// TIA Portal V21 export
// export: Created 2026-08-21T20:18:54.0096754Z, ExportSetting None, DisplayName Totally Integrated Automation Portal, DisplayVersion V21, DisplayName STEP 7 Professional, DisplayVersion V21, DisplayName STEP 7 Safety, DisplayVersion V21, DisplayName Tech WebApplication, DisplayVersion V21, DisplayName WinCC Basic/Comfort/Advanced, DisplayVersion V21, DisplayName WinCC Professional, DisplayVersion V21, DisplayName WinCC Unified, DisplayVersion V21
FUNCTION_BLOCK "MTPPIDCtrl_Type1"   // FB14, FBD
{ S7_Optimized_Access := 'TRUE' }
// stored: MemoryReserve 100, SetENOAutomatically false
   VAR_INPUT
      from_Actor { ExternalAccessible := 'False'; ExternalVisible := 'False'; ExternalWritable := 'False'} : "StruCm";
      SP_Ext { ExternalAccessible := 'False'; ExternalVisible := 'False'; ExternalWritable := 'False'} : Real;
      Service_Occupied { ExternalAccessible := 'False'; ExternalVisible := 'False'; ExternalWritable := 'False'} : Bool;
      Cmd_Auto { ExternalAccessible := 'False'; ExternalVisible := 'False'; ExternalWritable := 'False'} : Bool;
      Cmd_Man { ExternalAccessible := 'False'; ExternalVisible := 'False'; ExternalWritable := 'False'} : Bool;
      Cmd_SPExt { ExternalAccessible := 'False'; ExternalVisible := 'False'; ExternalWritable := 'False'} : Bool;
      Cmd_SPInt { ExternalAccessible := 'False'; ExternalVisible := 'False'; ExternalWritable := 'False'} : Bool;
      PV { ExternalAccessible := 'False'; ExternalVisible := 'False'; ExternalWritable := 'False'} : Word;
      PV_QB { ExternalAccessible := 'False'; ExternalVisible := 'False'; ExternalWritable := 'False'} : Bool := true;
      PV_Unit { ExternalAccessible := 'False'; ExternalVisible := 'False'; ExternalWritable := 'False'} : Int := 1342;
      Intlk04_In01 { ExternalAccessible := 'False'; ExternalVisible := 'False'; ExternalWritable := 'False'} : "DigVal";
      Intlk04_InvIn01 { ExternalAccessible := 'False'; ExternalVisible := 'False'; ExternalWritable := 'False'} : Bool;
      Intlk04_In1String : String;
      Intlk04_In02 { ExternalAccessible := 'False'; ExternalVisible := 'False'; ExternalWritable := 'False'} : "DigVal";
      Intlk04_InvIn02 { ExternalAccessible := 'False'; ExternalVisible := 'False'; ExternalWritable := 'False'} : Bool;
      Intlk04_In2String : String;
      Intlk04_In03 { ExternalAccessible := 'False'; ExternalVisible := 'False'; ExternalWritable := 'False'} : "DigVal";
      Intlk04_InvIn03 { ExternalAccessible := 'False'; ExternalVisible := 'False'; ExternalWritable := 'False'} : Bool;
      Intlk04_In3String : String;
      Intlk04_In04 { ExternalAccessible := 'False'; ExternalVisible := 'False'; ExternalWritable := 'False'} : "DigVal";
      Intlk04_InvIn04 { ExternalAccessible := 'False'; ExternalVisible := 'False'; ExternalWritable := 'False'} : Bool;
      Intlk04_In4String : String;
   END_VAR
   VAR_OUTPUT
      to_Actor { ExternalAccessible := 'False'; ExternalVisible := 'False'; ExternalWritable := 'False'} : "StruCm";
      Occupied { ExternalAccessible := 'False'; ExternalVisible := 'False'; ExternalWritable := 'False'} : Bool;   // Occupied by a Service procedure
      AutAct { ExternalAccessible := 'False'; ExternalVisible := 'False'; ExternalWritable := 'False'} : Bool;
      ManAct { ExternalAccessible := 'False'; ExternalVisible := 'False'; ExternalWritable := 'False'} : Bool;
      SP_ExtAct { ExternalAccessible := 'False'; ExternalVisible := 'False'; ExternalWritable := 'False'} : Bool;
      GrpErr { ExternalAccessible := 'False'; ExternalVisible := 'False'; ExternalWritable := 'False'} : Bool;
      PV_AH_Act { ExternalAccessible := 'False'; ExternalVisible := 'False'; ExternalWritable := 'False'} : Bool;
      PV_WH_Act { ExternalAccessible := 'False'; ExternalVisible := 'False'; ExternalWritable := 'False'} : Bool;
      PV_WL_Act { ExternalAccessible := 'False'; ExternalVisible := 'False'; ExternalWritable := 'False'} : Bool;
      PV_AL_Act { ExternalAccessible := 'False'; ExternalVisible := 'False'; ExternalWritable := 'False'} : Bool;
   END_VAR
   VAR
      AnIn_IDB { ExternalAccessible := 'False'; ExternalVisible := 'False'; ExternalWritable := 'False'} : "AnIn";
      Intlk04_IDB : "Intlk04";
      PIDConL_IDB { S7_SetPoint := 'True'} : "PIDConL";
      MTPPIDCtrl_IDB { ExternalVisible := 'False'; S7_SetPoint := 'True'} : "MTPPIDCtrl";
   END_VAR
   VAR_TEMP
      Intlock : "DigVal";
      PV_Out : "AnaVal";
      ScaleOut : "ScaVal";
      BadOut : "DigVal";
      CSF_NOP : "DigVal";
   END_VAR
   // Intlk04_In01.Value := true;
   // Intlk04_In02.Value := true;
   // Intlk04_In03.Value := true;
   // Intlk04_In04.Value := true;
BEGIN

REGION Network 1: Mod switch
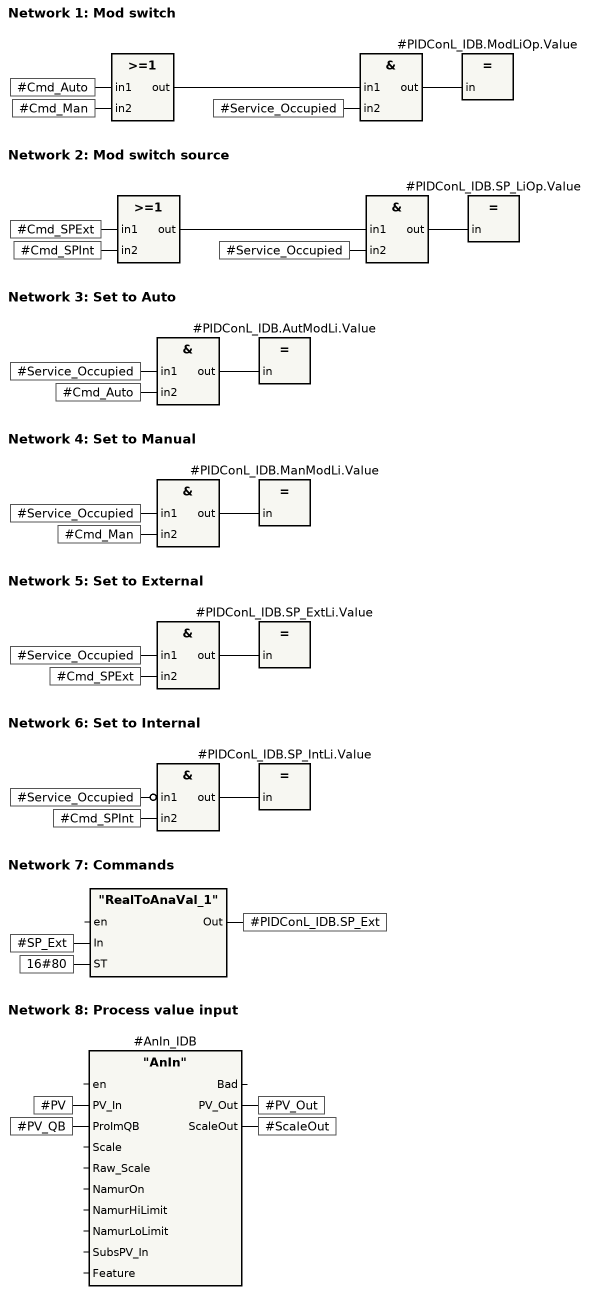
   #PIDConL_IDB.ModLiOp.Value := (#Cmd_Auto OR #Cmd_Man) AND #Service_Occupied;
END_REGION

REGION Network 2: Mod switch source
   #PIDConL_IDB.SP_LiOp.Value := (#Cmd_SPExt OR #Cmd_SPInt) AND #Service_Occupied;
END_REGION

REGION Network 3: Set to Auto
   #PIDConL_IDB.AutModLi.Value := #Service_Occupied AND #Cmd_Auto;
END_REGION

REGION Network 4: Set to Manual
   #PIDConL_IDB.ManModLi.Value := #Service_Occupied AND #Cmd_Man;
END_REGION

REGION Network 5: Set to External
   #PIDConL_IDB.SP_ExtLi.Value := #Service_Occupied AND #Cmd_SPExt;
END_REGION

REGION Network 6: Set to Internal
   #PIDConL_IDB.SP_IntLi.Value := NOT #Service_Occupied AND #Cmd_SPInt;
END_REGION

REGION Network 7: Commands
   "RealToAnaVal_1"(In := #SP_Ext, ST := 16#80, Out => #PIDConL_IDB.SP_Ext);
END_REGION

REGION Network 8: Process value input
   #AnIn_IDB(PV_In := #PV, ProImQB := #PV_QB, PV_Out => #PV_Out, ScaleOut => #ScaleOut);   // "AnIn"
END_REGION

REGION Network 9: CSF
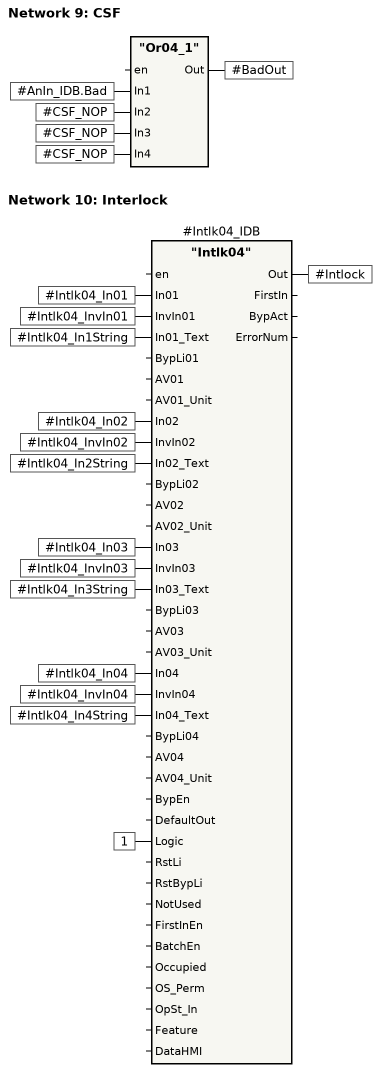
   "Or04_1"(In1 := #AnIn_IDB.Bad, In2 := #CSF_NOP, In3 := #CSF_NOP, In4 := #CSF_NOP, Out => #BadOut);
END_REGION

REGION Network 10: Interlock
   #Intlk04_IDB(In01 := #Intlk04_In01,   // "Intlk04"
                InvIn01 := #Intlk04_InvIn01,
                In01_Text := #Intlk04_In1String,
                In02 := #Intlk04_In02,
                InvIn02 := #Intlk04_InvIn02,
                In02_Text := #Intlk04_In2String,
                In03 := #Intlk04_In03,
                InvIn03 := #Intlk04_InvIn03,
                In03_Text := #Intlk04_In3String,
                In04 := #Intlk04_In04,
                InvIn04 := #Intlk04_InvIn04,
                In04_Text := #Intlk04_In4String,
                Logic := 1,
                Out => #Intlock);
END_REGION

REGION Network 11: PIDCtrL / PIDConL
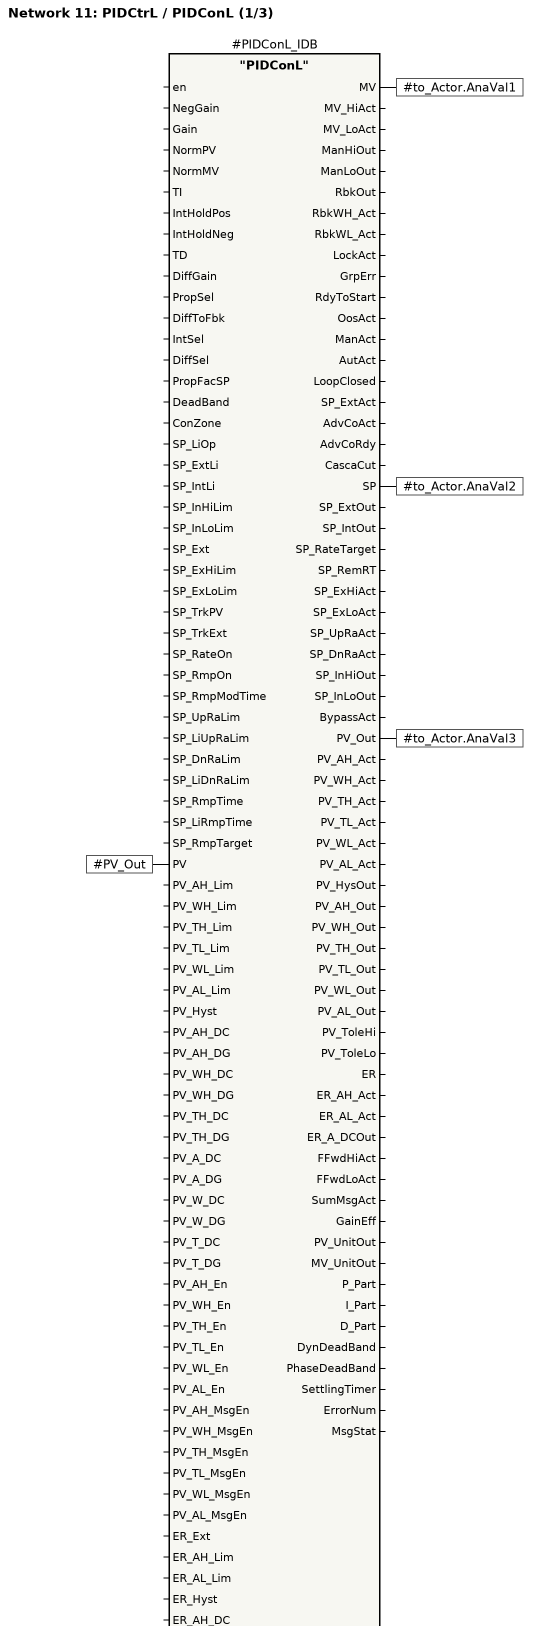
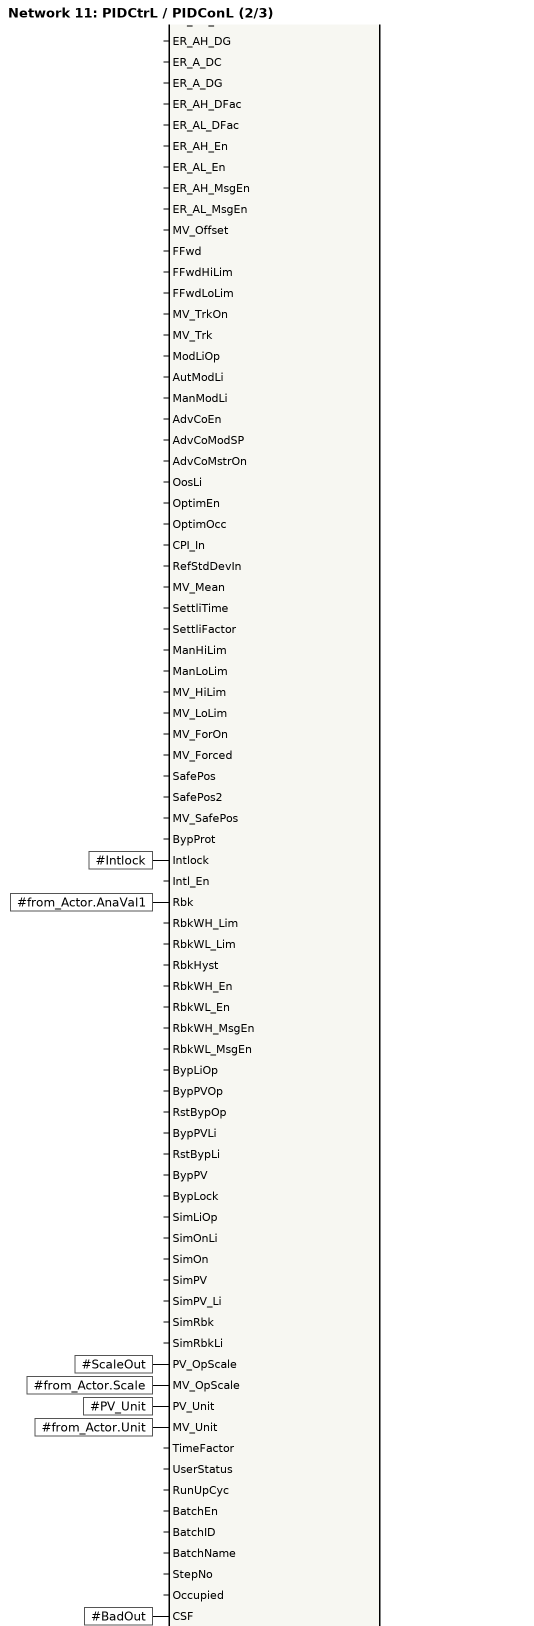
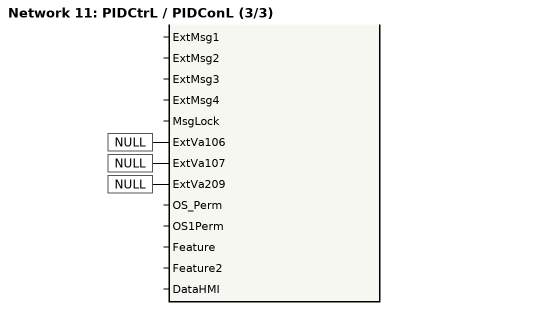
   #PIDConL_IDB(PV := #PV_Out,   // "PIDConL"
                Intlock := #Intlock,
                Rbk := #from_Actor.AnaVal1,
                PV_OpScale := #ScaleOut,
                MV_OpScale := #from_Actor.Scale,
                PV_Unit := #PV_Unit,
                MV_Unit := #from_Actor.Unit,
                CSF := #BadOut,
                ExtVa106 := NULL,
                ExtVa107 := NULL,
                ExtVa209 := NULL,
                MV => #to_Actor.AnaVal1,
                SP => #to_Actor.AnaVal2,
                PV_Out => #to_Actor.AnaVal3);
END_REGION

REGION Network 12: MTPPIDCtrl
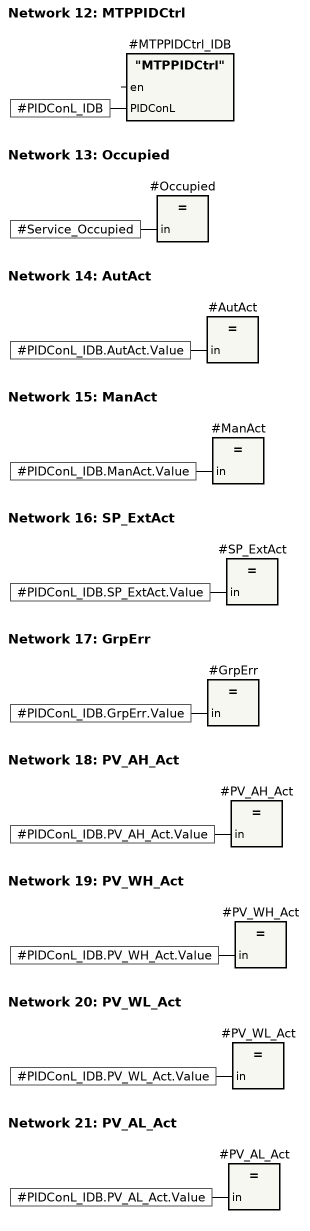
   #MTPPIDCtrl_IDB(PIDConL := #PIDConL_IDB);   // "MTPPIDCtrl"
END_REGION

REGION Network 13: Occupied
   #Occupied := #Service_Occupied;
END_REGION

REGION Network 14: AutAct
   #AutAct := #PIDConL_IDB.AutAct.Value;
END_REGION

REGION Network 15: ManAct
   #ManAct := #PIDConL_IDB.ManAct.Value;
END_REGION

REGION Network 16: SP_ExtAct
   #SP_ExtAct := #PIDConL_IDB.SP_ExtAct.Value;
END_REGION

REGION Network 17: GrpErr
   #GrpErr := #PIDConL_IDB.GrpErr.Value;
END_REGION

REGION Network 18: PV_AH_Act
   #PV_AH_Act := #PIDConL_IDB.PV_AH_Act.Value;
END_REGION

REGION Network 19: PV_WH_Act
   #PV_WH_Act := #PIDConL_IDB.PV_WH_Act.Value;
END_REGION

REGION Network 20: PV_WL_Act
   #PV_WL_Act := #PIDConL_IDB.PV_WL_Act.Value;
END_REGION

REGION Network 21: PV_AL_Act
   #PV_AL_Act := #PIDConL_IDB.PV_AL_Act.Value;
END_REGION
END_FUNCTION_BLOCK
